Fanuc KAREL source: kf00096.KL

-- PROVISIONAL review KL for V940-1; original PC SHA256 b30baa3b296a20c18f01224a1c9c619e86a10d90c6eb6c550e724f55c9e712b7
-- Incomplete behavior may be omitted. Consult companion uncertainty JSON. Do not deploy.
PROGRAM KF00096
%NOLOCKGROUP
BEGIN
  -- V9_ZERO_TABLE_METADATA_HINT layout=0002_ascii; no indexed target words; source/name/runtime held
  -- UNRESOLVED_PC offsets 5-16; opcodes 2E,23
  -- UNRESOLVED_PC offsets 21-32; opcodes 2E,23
  -- UNRESOLVED_PC offsets 37-67; opcodes 27,27,9D,22,22,22,22,31
  -- UNRESOLVED_PC offsets 72-76; opcodes 7F
END KF00096
